Staubli VAL3: getIFvalue.pgx

public program getIFvalue(string x_sKey, num x_nIndex, bool& x_bFinalResult)
  local num l_nSigType[3]
  local num l_i
  local num l_nSigValue[3]
  local bool l_bANDOR[2]
  local num l_nSigIndex[3]
  local bool l_bValue
  local bool l_bErr
  local bool l_bSetValue
  local num l_nResult[3]
  local bool l_bResult0[2]
  local num l_nValue
begin
  //l_nResult=0,null
  //         =1,true
  //         =2,false

  for l_i = 0 to 2
    l_nSigType[l_i]= trajTemp:tTrajItem[x_sKey].pPointItem[x_nIndex].pParaItem.iIfItem.nSigType[l_i]
    l_nSigValue[l_i]=trajTemp:tTrajItem[x_sKey].pPointItem[x_nIndex].pParaItem.iIfItem.nValue[l_i]
    l_nSigIndex[l_i]=trajTemp:tTrajItem[x_sKey].pPointItem[x_nIndex].pParaItem.iIfItem.nSigIndex[l_i]
  endFor
  l_bANDOR[0]=trajTemp:tTrajItem[x_sKey].pPointItem[x_nIndex].pParaItem.iIfItem.bANDOR[0]
  l_bANDOR[1]=trajTemp:tTrajItem[x_sKey].pPointItem[x_nIndex].pParaItem.iIfItem.bANDOR[1]

  for l_i = 0 to 2
    if l_nSigType[l_i]!=0 and l_nSigIndex[l_i]!=0
      switch l_nSigType[l_i]
        case 1
          //din
          call io:getDigIO(io:dInput[l_nSigIndex[l_i]],l_bValue,l_bErr)
          l_bSetValue=(l_nSigValue[l_i]!=0)
          if l_bSetValue==l_bValue
            l_nResult[l_i]=1
          else
            l_nResult[l_i]=2
          endIf
        break
        case 2
          //dout
          call io:getDigIO(io:dOutput[l_nSigIndex[l_i]],l_bValue,l_bErr)
          l_bSetValue=(l_nSigValue[l_i]!=0)
          if l_bSetValue==l_bValue
            l_nResult[l_i]=1
          else
            l_nResult[l_i]=2
          endIf
        break
        case 3
          //ain
          call io:getAnaIO(io:aInput[l_nSigIndex[l_i]],l_nValue,l_bErr)
          if l_nSigValue[l_i]==l_nValue
            l_nResult[l_i]=1
          else
            l_nResult[l_i]=2
          endIf
        break
        case 4
          //aout
          call io:getAnaIO(io:aOutput[l_nSigIndex[l_i]],l_nValue,l_bErr)
          if l_nSigValue[l_i]==l_nValue
            l_nResult[l_i]=1
          else
            l_nResult[l_i]=2
          endIf
        break
      endSwitch
    else
      l_nResult[l_i]=0
    endIf
  endFor

  //logic
 call logicIF(l_nResult[0],l_nResult[1],l_nResult[2],l_bANDOR[0],l_bANDOR[1],x_bFinalResult)

end
